Fanuc KAREL source: KA00057.KL

PROGRAM KA00057
%NOLOCKGROUP
VAR
  SRC: POSITION
  DST: VECTOR
BEGIN
  DST = SRC
END KA00057
